// FB RS and FB SR state codes.
{attribute 'qualified_only'}
{attribute 'to_string'}
TYPE
E_SafeLatchState :
(
    Undefined := 0,
    Stop := 2,
    Safe := 3,
    Set := 9
) BYTE;
END_TYPE

(* stored: Version 1.1.0.1
   DUT E_SafeLatchState: Id {929be28e-4d07-5c61-b708-4b9a648d47a5} *)
